Fanuc KAREL source: KT00042.KL

PROGRAM KT00042
%NOLOCKGROUP
VAR
  R1: REAL
  I2: INTEGER
  OUT: REAL
BEGIN
  R1 = 2.0
    I2 = 3
  OUT = R1 - I2
END KT00042
